// TIA Portal V21 export
FUNCTION_BLOCK "FB_AnaGlobalAccess"   // FB14, SCL
TITLE = Analyzer: global access inside an FB
{ S7_Optimized_Access := 'TRUE' }
// Rule C26g: a global DB and PLC tags are accessed inside the FB
// stored: MemoryReserve 100, SetENOAutomatically false
   VAR_OUTPUT
      Speed : Real;   // Speed setpoint from the global DB
   END_VAR
BEGIN

       #Speed := "DB_Machine".SpeedSetpoint;
       "ConveyorRun" := "StartButton";
END_FUNCTION_BLOCK
